(* IEC 61131-3 sources: SortJet_MasterSPS_Aufbau.fbsproj/07_Auftragsverwaltung/Job_Fremdanlage.prg.st^, 4 files *)

(* ---- Auftraege.act.st ---- *)
(* METADATA
{
	"v3Meta": {
		"objectGuid": "c249d517-2d16-45f2-b7bc-658c62d8cf35"
	}
}
*)
ACTION Auftraege
//-------------------------------------------------------------------------------------------------
// AUFTRAG: M_SB0_MMI_ISOQUITTUNG
//-------------------------------------------------------------------------------------------------
(* Hinweis:
   - Unabhaengige Quittung der Sondergläser durch Tasterdruck anfordern
*)
IF ( M_SB0_MMI_ISOQUITTUNG ) THEN
  M_SB0_MMI_ISOQUITTUNG:=FALSE;

  CASE tMmi2SpsInfo.wISOStation OF

    cERSTE_FREMDANLAGE..cLETZTE_FREMDANLAGE:
      aSchnittstelleAuslauf[tMmi2SpsInfo.wISOStation].wpAuftragsTyp := tMmi2SpsInfo.wISOAuftragsID;
      aSchnittstelleAuslauf[tMmi2SpsInfo.wISOStation].bpStarteIGEvent := TRUE;

  END_CASE

END_IF

//-------------------------------------------------------------------------------------------------
// AUFTRAG: M_SB0_MMI_SORTIERUNGCANCELISOLINEEVENT
//-------------------------------------------------------------------------------------------------
(* Hinweis:
   -  Abbruch des offenen ISO Line Events
*)

IF ( M_SB0_MMI_SORTIERUNGCANCELISOLINEEVENT ) THEN
  M_SB0_MMI_SORTIERUNGCANCELISOLINEEVENT := FALSE;

  CASE tMmi2SpsInfo.wDeleteISOLinienStationNr OF

    cERSTE_FREMDANLAGE..cLETZTE_FREMDANLAGE:
      aSchnittstelleAuslauf[tMmi2SpsInfo.wDeleteISOLinienStationNr].bpResetISOLinieEvent := TRUE;

  END_CASE

END_IF

//-------------------------------------------------------------------------------------------------
// AUFTRAG: M_SB0_MMI_AUFTRAGSDATEN_FREMDANLAGE
//-------------------------------------------------------------------------------------------------
(* Hinweis:
   -  Auftragsdaten fuer die Fremdanlage
*)
IF ( M_SB0_MMI_AUFTRAGSDATEN_FREMDANLAGE ) THEN
  M_SB0_MMI_AUFTRAGSDATEN_FREMDANLAGE := FALSE;

  CASE tMmi2SpsInfo.wFremdanlageNr OF

    cERSTE_FREMDANLAGE..cLETZTE_FREMDANLAGE:
      (* Hinweis:
         - Es folgt hier keine weitere Nachricht
      *)
      IF ( tMmi2SpsInfo.wNachrichtenAnzahl = 1 ) THEN
        stAuftragScheibenIDs.adwScheibenID_1 := ScheibenID(tMmi2SpsInfo.wFremdanlageNr, tMmi2SpsInfo.adwScheibenID_1);
        stAuftragScheibenIDs.adwScheibenID_2 := ScheibenID(tMmi2SpsInfo.wFremdanlageNr, tMmi2SpsInfo.adwScheibenID_2);
        stAuftragScheibenIDs.adwScheibenID_3 := ScheibenID(tMmi2SpsInfo.wFremdanlageNr, tMmi2SpsInfo.adwScheibenID_3);
        stAuftragScheibenIDs.adwScheibenID_4 := ScheibenID(tMmi2SpsInfo.wFremdanlageNr, tMmi2SpsInfo.adwScheibenID_4);

        aSchnittstelleAuslauf[tMmi2SpsInfo.wFremdanlageNr].AuftragsSpeicher.ppEingabeWert.wScheibenAnzahl := tMmi2SpsInfo.wScheibenanzahl;
        aSchnittstelleAuslauf[tMmi2SpsInfo.wFremdanlageNr].AuftragsSpeicher.ppEingabeWert.stScheibenID    := stAuftragScheibenIDs;
        aSchnittstelleAuslauf[tMmi2SpsInfo.wFremdanlageNr].AuftragsSpeicher( bpWerteSchreiben  := TRUE );

        stAuftragScheibenIDs.adwScheibenID_1[0]  := 0;
        stAuftragScheibenIDs.adwScheibenID_1[1]  := 0;
        stAuftragScheibenIDs.adwScheibenID_1[2]  := 0;
        stAuftragScheibenIDs.adwScheibenID_1[3]  := 0;
        stAuftragScheibenIDs.adwScheibenID_2[0]  := 0;
        stAuftragScheibenIDs.adwScheibenID_2[1]  := 0;
        stAuftragScheibenIDs.adwScheibenID_2[2]  := 0;
        stAuftragScheibenIDs.adwScheibenID_2[3]  := 0;
        stAuftragScheibenIDs.adwScheibenID_3[0]  := 0;
        stAuftragScheibenIDs.adwScheibenID_3[1]  := 0;
        stAuftragScheibenIDs.adwScheibenID_3[2]  := 0;
        stAuftragScheibenIDs.adwScheibenID_3[3]  := 0;
        stAuftragScheibenIDs.adwScheibenID_4[0]  := 0;
        stAuftragScheibenIDs.adwScheibenID_4[1]  := 0;
        stAuftragScheibenIDs.adwScheibenID_4[2]  := 0;
        stAuftragScheibenIDs.adwScheibenID_4[3]  := 0;
        stAuftragScheibenIDs.adwScheibenID_5[0]  := 0;
        stAuftragScheibenIDs.adwScheibenID_5[1]  := 0;
        stAuftragScheibenIDs.adwScheibenID_5[2]  := 0;
        stAuftragScheibenIDs.adwScheibenID_5[3]  := 0;
        stAuftragScheibenIDs.adwScheibenID_6[0]  := 0;
        stAuftragScheibenIDs.adwScheibenID_6[1]  := 0;
        stAuftragScheibenIDs.adwScheibenID_6[2]  := 0;
        stAuftragScheibenIDs.adwScheibenID_6[3]  := 0;

      (* Hinweis:
         - Es muss nicht noch auf eine Nachricht gewartet werden
      *)
      ELSE

        blUeberwachungFolgeNachricht := TRUE;

        CASE tMmi2SpsInfo.wNachrichtenIndex OF

          cNACHRICHTEN_INDEX_1:
            ablNachrichtEmpfangen[1] := TRUE;

            stAuftragScheibenIDs.adwScheibenID_1 := ScheibenID(tMmi2SpsInfo.wFremdanlageNr, tMmi2SpsInfo.adwScheibenID_1);
            stAuftragScheibenIDs.adwScheibenID_2 := ScheibenID(tMmi2SpsInfo.wFremdanlageNr, tMmi2SpsInfo.adwScheibenID_2);
            stAuftragScheibenIDs.adwScheibenID_3 := ScheibenID(tMmi2SpsInfo.wFremdanlageNr, tMmi2SpsInfo.adwScheibenID_3);
            stAuftragScheibenIDs.adwScheibenID_4 := ScheibenID(tMmi2SpsInfo.wFremdanlageNr, tMmi2SpsInfo.adwScheibenID_4);

          cNACHRICHTEN_INDEX_2:
            ablNachrichtEmpfangen[2] := TRUE;

            // Zweite Nachricht: Scheiben-ID 1 und 2 enthalten die Scheiben 5 und 6
            stAuftragScheibenIDs.adwScheibenID_5 := ScheibenID(tMmi2SpsInfo.wFremdanlageNr, tMmi2SpsInfo.adwScheibenID_1);
            stAuftragScheibenIDs.adwScheibenID_6 := ScheibenID(tMmi2SpsInfo.wFremdanlageNr, tMmi2SpsInfo.adwScheibenID_2);

          ELSE
            wpgFehlerdaten[0] := tMmi2SpsInfo.wNachrichtenIndex;
            SpsWarnung( eFehler_Schnittstelle,
                        cMELDUNG_SCHNITTSTELLE_AUFTRAGSDATEN_SCHNITTSTELLE_NACHRICHTENINDEX_FEHLERHAFT,
                        tMmi2SpsInfo.wNachrichtenIndex,
                        AutomatikkreisBestimmen(0),
                        wpgFehlerdaten );

        END_CASE

        (* Hinweis:
           - Werte zuruecksetzen wenn alle Nachrichten Empfangen worden sind
        *)
        IF (  ablNachrichtEmpfangen[1]
             AND ablNachrichtEmpfangen[2] )
        THEN
          aSchnittstelleAuslauf[tMmi2SpsInfo.wFremdanlageNr].AuftragsSpeicher.ppEingabeWert.stScheibenID    := stAuftragScheibenIDs;
          aSchnittstelleAuslauf[tMmi2SpsInfo.wFremdanlageNr].AuftragsSpeicher.ppEingabeWert.wScheibenAnzahl := tMmi2SpsInfo.wScheibenanzahl;
          aSchnittstelleAuslauf[tMmi2SpsInfo.wFremdanlageNr].AuftragsSpeicher( bpWerteSchreiben  := TRUE );

          stAuftragScheibenIDs.adwScheibenID_1[0]  := 0;
          stAuftragScheibenIDs.adwScheibenID_1[1]  := 0;
          stAuftragScheibenIDs.adwScheibenID_1[2]  := 0;
          stAuftragScheibenIDs.adwScheibenID_1[3]  := 0;
          stAuftragScheibenIDs.adwScheibenID_2[0]  := 0;
          stAuftragScheibenIDs.adwScheibenID_2[1]  := 0;
          stAuftragScheibenIDs.adwScheibenID_2[2]  := 0;
          stAuftragScheibenIDs.adwScheibenID_2[3]  := 0;
          stAuftragScheibenIDs.adwScheibenID_3[0]  := 0;
          stAuftragScheibenIDs.adwScheibenID_3[1]  := 0;
          stAuftragScheibenIDs.adwScheibenID_3[2]  := 0;
          stAuftragScheibenIDs.adwScheibenID_3[3]  := 0;
          stAuftragScheibenIDs.adwScheibenID_4[0]  := 0;
          stAuftragScheibenIDs.adwScheibenID_4[1]  := 0;
          stAuftragScheibenIDs.adwScheibenID_4[2]  := 0;
          stAuftragScheibenIDs.adwScheibenID_4[3]  := 0;
          stAuftragScheibenIDs.adwScheibenID_5[0]  := 0;
          stAuftragScheibenIDs.adwScheibenID_5[1]  := 0;
          stAuftragScheibenIDs.adwScheibenID_5[2]  := 0;
          stAuftragScheibenIDs.adwScheibenID_5[3]  := 0;
          stAuftragScheibenIDs.adwScheibenID_6[0]  := 0;
          stAuftragScheibenIDs.adwScheibenID_6[1]  := 0;
          stAuftragScheibenIDs.adwScheibenID_6[2]  := 0;
          stAuftragScheibenIDs.adwScheibenID_6[3]  := 0;

          ablNachrichtEmpfangen[1]     := FALSE;
          ablNachrichtEmpfangen[2]     := FALSE;
          blUeberwachungFolgeNachricht := FALSE;

        END_IF

      END_IF

    ELSE
      ;

  END_CASE

END_IF
END_ACTION

(* ---- Fremdanlage.meth.st ---- *)
(* METADATA
{
	"v3Meta": {
		"objectGuid": "cf66fcf2-cc11-47d6-b197-d71c762428b0"
	}
}
*)
METHOD INTERNAL Fremdanlage
VAR_INPUT
  wFremdanlage                  : WORD;
  wVorgaenger                   : WORD;
  wAutomatikkreis               : WORD;
  bDurchtransportierendeStation : BOOL;
END_VAR
VAR
  ptSender                    : REFERENCE TO StationBasisParameter_ST;
  ptAuftragsdatenSender       : REFERENCE TO Auftragsdaten_ST;
  ptAuftragsdatenVorgaenger   : REFERENCE TO Auftragsdaten_ST;
END_VAR

// Hinweis:
// - Glas-Sender ist die Transferstation 1 des Fremdanlagen-Auftrags (Shuttle, Transfershuttle oder Station)
// - Shuttle und Transfershuttle (MK bStationIstShuttle) legen den Auftrag der Fremdanlage selbst an
// - Bei einer Station legt die Fremdanlage den Austransport-Auftrag ihres Vorgaengers an
ptSender              REF= getBasis( AuftragsdatenFremdanlage[wFremdanlage].wTransferstationsNr1 );
ptAuftragsdatenSender REF= getAuftragsdaten( AuftragsdatenFremdanlage[wFremdanlage].wTransferstationsNr1,
                                             AuftragsdatenFremdanlage[wFremdanlage].wTransferwand );
ptAuftragsdatenVorgaenger REF= getAuftragsdaten( wVorgaenger, cWAND_1 );

//-------------------------------------------------------------------------------------------------
// STEUERUNG EINTRANSPORT
//-------------------------------------------------------------------------------------------------
IF ( AuftragsdatenFremdanlage[wFremdanlage].wAuftrag = eStation_Eintransport ) THEN
  CASE astplEintransportFremdanlage[wFremdanlage] OF
    // EINTRANSPORT ===========================================
    STEP_0_E:
      (* Hinweis:
         - Ueberpruefung des Sicherheitskreises
      *)
      astplEintransportFremdanlage[wFremdanlage] := STEP_10_E;

    // EINTRANSPORT ===========================================
    STEP_10_E:
      // ---------------------------------------------------------------------------------------
      // GLAS-SENDER PRUEFUNG
      //
      //  Hinweis:
      // - n/c
      // ---------------------------------------------------------------------------------------

      (* Hinweis:
         - Glas- Sender bestimmen und merken
      *)
      IF (     __ISVALIDREF( ptSender )
           AND_THEN __ISVALIDREF( ptSender.stMKs )
           AND_THEN ptSender.stMKs.stSchnittstellendaten.bStationIstShuttle )
      THEN
        starrFremdanlageAuslaufStationBasisParameter[AuftragsdatenFremdanlage[wFremdanlage].wStationsNr].InGlasTransportVorgaenger[cWAND_1] := ptSender.OutGlasTransport[AuftragsdatenFremdanlage[wFremdanlage].wTransferwand];
        astplEintransportFremdanlage[wFremdanlage] := STEP_40_E;
      ELSE
        astplEintransportFremdanlage[wFremdanlage] := STEP_30_E;
      END_IF

    // EINTRANSPORT ===========================================
    STEP_30_E:
      // ---------------------------------------------------------------------------------------
      // PRUEFUNG AUFTRAGSSTATUS GLAS-SENDER
      //
      //  Hinweis:
      // - n/c
      // ---------------------------------------------------------------------------------------
      IF ( __ISVALIDREF( ptAuftragsdatenVorgaenger ) ) THEN

        IF ( ( ptAuftragsdatenVorgaenger.wAuftrag = eStation_Belegt )
             OR ( ptAuftragsdatenVorgaenger.wAuftrag = eStation_Warte_Auf_Austransport ) )
           OR ( ( ptAuftragsdatenVorgaenger.wAuftrag = eStation_Kein_Auftrag ) AND bDurchtransportierendeStation )
        THEN

          IF bDurchtransportierendeStation THEN
            ptAuftragsdatenVorgaenger := AuftragsdatenUmkopieren(FALSE, TRUE, AuftragsdatenFremdanlage[wFremdanlage]);
            ptAuftragsdatenVorgaenger.wAuftrag := eStation_Durchtransport;
          ELSE
            ptAuftragsdatenVorgaenger := AuftragsdatenUmkopieren(FALSE, FALSE, AuftragsdatenFremdanlage[wFremdanlage]);
            ptAuftragsdatenVorgaenger.wAuftrag := eStation_Austransport;
          END_IF

          astplEintransportFremdanlage[wFremdanlage] := STEP_40_E;

        END_IF

      END_IF

    // EINTRANSPORT ===========================================
    STEP_40_E:
      (* Hinweis:
         - Abgeschlossen, sobald der Glas-Sender seinen Austransport (bzw. Durchtransport) beendet hat
      *)
      IF bDurchtransportierendeStation THEN
        IF ( NOT __ISVALIDREF( ptAuftragsdatenVorgaenger ) ) OR_ELSE ( ptAuftragsdatenVorgaenger.wAuftrag <> eStation_Durchtransport ) THEN
          astplEintransportFremdanlage[wFremdanlage] := STEP_1000_E;
        END_IF
      ELSE
        IF ( NOT __ISVALIDREF( ptAuftragsdatenSender ) ) OR_ELSE ( ptAuftragsdatenSender.wAuftrag <> eStation_Austransport ) THEN
          astplEintransportFremdanlage[wFremdanlage] := STEP_1000_E;
        END_IF
      END_IF

    // EINTRANSPORT ===========================================
    STEP_900_E:
      abpFehler[wAutomatikkreis] := TRUE;

    // EINTRANSPORT ===========================================
    STEP_1000_E:
      AuftragsdatenFremdanlage[wFremdanlage].wAuftrag := eStation_Kein_Auftrag;

  // EINTRANSPORT ===========================================
  END_CASE
END_IF

IF ( NOT (AuftragsdatenFremdanlage[wFremdanlage].wAuftrag = eStation_Eintransport) ) THEN

  IF ( astplEintransportFremdanlage[wFremdanlage] > STEP_0_E ) THEN
    astplEintransportFremdanlage[wFremdanlage] := STEP_0_E;
  END_IF

END_IF
END_METHOD

(* ---- Reset.act.st ---- *)
(* METADATA
{
	"v3Meta": {
		"objectGuid": "ba21d831-07aa-4eb0-a98f-ca51ada32f1d"
	}
}
*)
ACTION Reset
//-------------------------------------------------------------------------------------------------
// AKTION: RESET
//-------------------------------------------------------------------------------------------------

FOR wlIndexReset := cERSTER_AUTOMATIKKREIS TO cLETZTER_AUTOMATIKKREIS DO

  IF ( abpReset[wlIndexReset] ) THEN

    ablNachrichtEmpfangen[1]     := FALSE;
    ablNachrichtEmpfangen[2]     := FALSE;
    blUeberwachungFolgeNachricht := FALSE;
    abpReset[wlIndexReset]       := FALSE;

    // Schnittstelle Auslauf Reset
    FOR wlIndex := cERSTE_FREMDANLAGE_AUSLAUF TO cLETZTE_FREMDANLAGE_AUSLAUF DO
      IF StationInAutomatikkreis(starrFremdanlageAuslaufStationBasisParameter[wlIndex].stMKs.eaAutomatikkreis, wlIndexReset) THEN
        AuftragsdatenFremdanlage[wlIndex].wAuftrag := eStation_Kein_Auftrag;
        starrFremdanlageAuslaufStationBasisParameter[wlIndex].bReset := NOT starrFremdanlageAuslaufStationBasisParameter[wlIndex].stMKs.bDeaktivieren;
      END_IF
    END_FOR

    // Schnittstelle Einlauf Reset
    FOR wlIndex := cERSTE_FREMDANLAGE_EINLAUF TO cLETZTE_FREMDANLAGE_EINLAUF DO
      IF StationInAutomatikkreis(starrFremdanlageEinlaufStationBasisParameter[wlIndex].stMKs.eaAutomatikkreis, wlIndexReset) THEN
        AuftragsdatenFremdanlage[wlIndex].wAuftrag := eStation_Kein_Auftrag;
        starrFremdanlageEinlaufStationBasisParameter[wlIndex].bReset := NOT starrFremdanlageEinlaufStationBasisParameter[wlIndex].stMKs.bDeaktivieren;
      END_IF
    END_FOR

  END_IF

END_FOR
END_ACTION

(* ---- ScheibenID.meth.st ---- *)
(* METADATA
{
	"v3Meta": {
		"objectGuid": "e658493f-ee55-49d1-b74f-ae85f8ce4fd2"
	}
}
*)
METHOD PRIVATE ScheibenID : ARRAY [0..3] OF DWORD
VAR_INPUT
  wFremdanlage  : WORD;
  adwScheibenID : ARRAY [0..3] OF DWORD;
END_VAR

// Hinweis:
// - Scheiben-ID aus dem MMI uebernehmen, ETX nur entfernen wenn per MK aktiviert (stFremdanlage.bRemoveETX)
IF ( starrFremdanlageAuslaufStationBasisParameter[wFremdanlage].stMKs.stFremdanlage.bRemoveETX ) THEN
  ScheibenID := RemoveETX( adwScheibenID );
ELSE
  ScheibenID := adwScheibenID;
END_IF
END_METHOD
